// TIA Portal V15.1 export
// export: Created 2026-11-11T00:40:31.1045989Z, ExportSetting WithDefaults, DisplayName Totally Integrated Automation Portal, DisplayVersion V15.1, DisplayName TIA Portal Openness, DisplayVersion V15.1, DisplayName STEP 7 Professional, DisplayVersion V15.1, DisplayName WinCC Professional, DisplayVersion V15.1
Screen "Alarms"  480x272, Number=5, Template=Template_1
  ScreenLayer 
    Rectangle "Panel_Panel" at 0,0 size 480x26
    TextField "Text_LCP_01_Alarms" at 6,2 size 300x22  Text="LCP-01 Alarms"
    TextField "Text_E_STOP_RESET_Sys_Alm_EStop" at 330,3 size 146x20  Text="E-STOP / RESET"
      SingleBitVisibilityAnimation "VisibilityAnimation"
        tag Sys_Alm_EStop
    Button "Nav_Root_screen" at 2,236 size 76x34  Mode=Text, TextOff="Overview", TextOn="Overview"
      on Press: ActivateScreen(Screen name := Root screen, Object number := 0)
    Button "Nav_BR01" at 82,236 size 76x34  Mode=Text, TextOff="BR01", TextOn="BR01"
      on Press: ActivateScreen(Screen name := BR01, Object number := 0)
    Button "Nav_BR02" at 162,236 size 76x34  Mode=Text, TextOff="BR02", TextOn="BR02"
      on Press: ActivateScreen(Screen name := BR02, Object number := 0)
    Button "Nav_Scrubber" at 242,236 size 76x34  Mode=Text, TextOff="Scrubber", TextOn="Scrubber"
      on Press: ActivateScreen(Screen name := Scrubber, Object number := 0)
    Button "Nav_Alarms" at 322,236 size 76x34  Mode=Text, TextOff="Alarms", TextOn="Alarms"
      on Press: ActivateScreen(Screen name := , Object number := 0)
    Button "Nav_Settings" at 402,236 size 76x34  Mode=Text, TextOff="Settings", TextOn="Settings"
      on Press: ActivateScreen(Screen name := Settings, Object number := 0)
    Rectangle "Panel_Alarm_list" at 4,30 size 472x202
